(* IEC 61131-3 sources: s7-to-codesys/src/POUs/S7Compat/F_S7TimeDiff, 1 file *)

(* ---- F_S7TimeDiff.decl.st ---- *)
// Назначение: прошедшее время между моментами tStart и tNow (оба — F_S7Now) для ST-двойника S7-GRAPH: время
//             активности шага Si.T. Разность — по модулю 2^32 мс: переход TIME через ноль (около 49,7 суток
//             работы ПЛК) не даёт отрицательного или огромного значения, пока шаг активен меньше 2^32 мс.
// Автор:      kr0nsch
// Версия:     1.2.0
// Документ:   docs/MAPPING_GRAPH.md; docs/ASSUMPTIONS.md, запись L18
FUNCTION F_S7TimeDiff : TIME
VAR_INPUT
    tNow : TIME;    // текущий момент (F_S7Now)
    tStart : TIME;  // момент активации шага (F_S7Now)
END_VAR
